Fanuc KAREL source: KB00108.KL

PROGRAM KB00108
%NOLOCKGROUP
%ENVIRONMENT PBQMGR
VAR
  P1: INTEGER
  P2: INTEGER
  P3: QUEUE_TYPE
  P4: ARRAY[4] OF INTEGER
  P5: INTEGER
BEGIN
  P1 = 1
  P2 = 1
  P4[1] = 1
  P5 = 1
  INSERT_QUEUE(P1, P2, P3, P4, P5)
END KB00108
